ABB RAPID module: CalibData.modx

MODULE CalibData
    PERS tooldata EE_tool:=[TRUE,[[0,0,70],[1,0,0,0]],[1,[0,0,1],[1,0,0,0],0,0,0]];
ENDMODULE
